Fanuc KAREL source: KS00020.KL

PROGRAM KS00020
%NOLOCKGROUP
TYPE
  REC_T = STRUCTURE
    VALUE: INTEGER
    FLAG: BOOLEAN
  ENDSTRUCTURE
VAR
  A: FILE
  B: FILE
  FLAG: BOOLEAN
  N: INTEGER
  STATUS: INTEGER
  PN: STRING[80]
  VN: STRING[80]
BEGIN
  PN = ''
  VN = 'A'
  GET_VAR(N, PN, VN, A, STATUS)
END KS00020
